ABB RAPID module: Module1_backup.mod

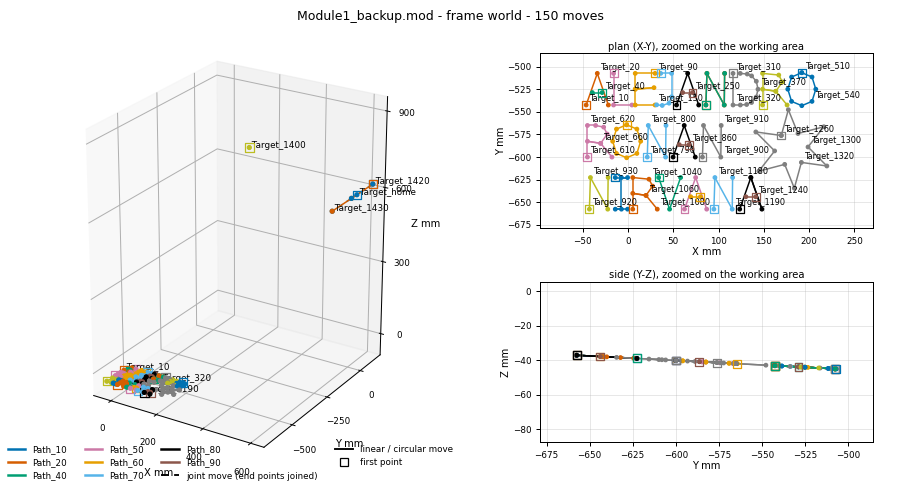
[picture p0: tool path of Module1_backup.mod in frame world, 150 of 178 moves have a stored position in this frame; points joined in program order, loops and branches not executed]
MODULE Module1
    PERS tooldata TOOLLAB1:=[TRUE,[[-6.48,-1.157,131.856],[0.965925826,0,0.258819045,0]],[1,[0,0,1],[1,0,0,0],0,0,0]];
    TASK PERS wobjdata Workobject_4:=[FALSE,TRUE,"",[[-82.07,-709.823595625,-134.482953476],[0.018509898,0.706864473,0.706864473,-0.018509898]],[[0,0,-100],[1,0,0,0]]];
    CONST robtarget Target_10:=[[162.356,35.679,0],[1,0,0,0],[-2,-1,0,1],[9E+09,9E+09,9E+09,9E+09,9E+09,9E+09]];
    CONST robtarget Target_20:=[[197.357,47.989,0],[1,0,0,0],[-2,-1,0,1],[9E+09,9E+09,9E+09,9E+09,9E+09,9E+09]];
    CONST robtarget Target_30:=[[162.356,60.2,0],[1,0,0,0],[-2,-1,0,1],[9E+09,9E+09,9E+09,9E+09,9E+09,9E+09]];
    CONST robtarget Target_40:=[[176.113,53.293,0],[1,0,0,0],[-2,-1,0,1],[9E+09,9E+09,9E+09,9E+09,9E+09,9E+09]];
    CONST robtarget Target_50:=[[176.113,42.487,0],[1,0,0,0],[-2,-1,0,1],[9E+09,9E+09,9E+09,9E+09,9E+09,9E+09]];
    VAR robtarget lift:=[[176.113,42.487,0],[0.707106781,0,0,-0.707106781],[-2,-1,0,1],[9E+09,9E+09,9E+09,9E+09,9E+09,9E+09]];
    CONST robtarget Target_60:=[[197.357,65.972,0],[1,0,0,0],[-2,-1,0,1],[9E+09,9E+09,9E+09,9E+09,9E+09,9E+09]];
    CONST robtarget Target_70:=[[162.356,65.972,0],[1,0,0,0],[-2,-1,0,1],[9E+09,9E+09,9E+09,9E+09,9E+09,9E+09]];
    CONST robtarget Target_80:=[[162.356,86.252,0],[1,0,0,0],[-2,-1,0,1],[9E+09,9E+09,9E+09,9E+09,9E+09,9E+09]];
    CONST robtarget Target_90:=[[197.357,111.808,0],[1,0,0,0],[-2,-1,0,1],[9E+09,9E+09,9E+09,9E+09,9E+09,9E+09]];
    CONST robtarget Target_100:=[[197.357,89.911,0],[1,0,0,0],[-2,-1,0,1],[9E+09,9E+09,9E+09,9E+09,9E+09,9E+09]];
    CONST robtarget Target_110:=[[179.857,89.911,0],[1,0,0,0],[-2,-1,0,1],[9E+09,9E+09,9E+09,9E+09,9E+09,9E+09]];
    CONST robtarget Target_120:=[[181.559,110.645,0],[1,0,0,0],[-2,-1,0,1],[9E+09,9E+09,9E+09,9E+09,9E+09,9E+09]];
    CONST robtarget Target_130:=[[179.857,89.911,0],[1,0,0,0],[-2,-1,0,1],[9E+09,9E+09,9E+09,9E+09,9E+09,9E+09]];
    CONST robtarget Target_140:=[[162.356,89.911,0],[1,0,0,0],[-2,-1,0,1],[9E+09,9E+09,9E+09,9E+09,9E+09,9E+09]];
    CONST robtarget Target_150:=[[162.356,111.808,0],[1,0,0,0],[-2,-1,0,1],[9E+09,9E+09,9E+09,9E+09,9E+09,9E+09]];
    CONST robtarget Target_160:=[[197.357,118.048,0],[1,0,0,0],[-2,-1,0,1],[9E+09,9E+09,9E+09,9E+09,9E+09,9E+09]];
    CONST robtarget Target_170:=[[197.357,130.103,0],[1,0,0,0],[-2,-1,0,1],[9E+09,9E+09,9E+09,9E+09,9E+09,9E+09]];
    CONST robtarget Target_180:=[[171.461,130.103,0],[1,0,0,0],[-2,-1,0,1],[9E+09,9E+09,9E+09,9E+09,9E+09,9E+09]];
    CONST robtarget Target_190:=[[164.37,127.295,0],[1,0,0,0],[-2,-1,0,1],[9E+09,9E+09,9E+09,9E+09,9E+09,9E+09]];
    CONST robtarget Target_200:=[[161.874,119.75,0],[1,0,0,0],[-2,-1,0,1],[9E+09,9E+09,9E+09,9E+09,9E+09,9E+09]];
    CONST robtarget Target_210:=[[162.555,113.567,0],[1,0,0,0],[-2,-1,0,1],[9E+09,9E+09,9E+09,9E+09,9E+09,9E+09]];
    CONST robtarget Target_220:=[[162.356,135.549,0],[1,0,0,0],[-2,-1,0,1],[9E+09,9E+09,9E+09,9E+09,9E+09,9E+09]];
    CONST robtarget Target_230:=[[197.357,147.859,0],[1,0,0,0],[-2,-1,0,1],[9E+09,9E+09,9E+09,9E+09,9E+09,9E+09]];
    CONST robtarget Target_240:=[[162.356,160.07,0],[1,0,0,0],[-2,-1,0,1],[9E+09,9E+09,9E+09,9E+09,9E+09,9E+09]];
    CONST robtarget Target_250:=[[176.113,153.163,0],[1,0,0,0],[-2,-1,0,1],[9E+09,9E+09,9E+09,9E+09,9E+09,9E+09]];
    CONST robtarget Target_260:=[[176.113,142.356,0],[1,0,0,0],[-2,-1,0,1],[9E+09,9E+09,9E+09,9E+09,9E+09,9E+09]];
    CONST robtarget Target_310:=[[197.357,197.978,0],[1,0,0,0],[-2,-1,0,1],[9E+09,9E+09,9E+09,9E+09,9E+09,9E+09]];
    CONST robtarget Target_320:=[[162.356,197.978,0],[1,0,0,0],[-2,-1,0,1],[9E+09,9E+09,9E+09,9E+09,9E+09,9E+09]];
    CONST robtarget Target_330:=[[162.356,206.033,0],[1,0,0,0],[-2,-1,0,1],[9E+09,9E+09,9E+09,9E+09,9E+09,9E+09]];
    CONST robtarget Target_340:=[[162.924,213.025,0],[1,0,0,0],[-2,-1,0,1],[9E+09,9E+09,9E+09,9E+09,9E+09,9E+09]];
    CONST robtarget Target_350:=[[165.164,218.429,0],[1,0,0,0],[-2,-1,0,1],[9E+09,9E+09,9E+09,9E+09,9E+09,9E+09]];
    CONST robtarget Target_360:=[[171.177,223.633,0],[1,0,0,0],[-2,-1,0,1],[9E+09,9E+09,9E+09,9E+09,9E+09,9E+09]];
    CONST robtarget Target_370:=[[179.829,225.576,0],[1,0,0,0],[-2,-1,0,1],[9E+09,9E+09,9E+09,9E+09,9E+09,9E+09]];
    CONST robtarget Target_380:=[[188.636,223.718,0],[1,0,0,0],[-2,-1,0,1],[9E+09,9E+09,9E+09,9E+09,9E+09,9E+09]];
    CONST robtarget Target_390:=[[194.578,218.485,0],[1,0,0,0],[-2,-1,0,1],[9E+09,9E+09,9E+09,9E+09,9E+09,9E+09]];
    CONST robtarget Target_400:=[[196.62,213.692,0],[1,0,0,0],[-2,-1,0,1],[9E+09,9E+09,9E+09,9E+09,9E+09,9E+09]];
    CONST robtarget Target_410:=[[197.357,205.948,0],[1,0,0,0],[-2,-1,0,1],[9E+09,9E+09,9E+09,9E+09,9E+09,9E+09]];
    CONST robtarget Target_420:=[[162.356,230.625,0],[1,0,0,0],[-2,-1,0,1],[9E+09,9E+09,9E+09,9E+09,9E+09,9E+09]];
    CONST robtarget Target_430:=[[197.357,230.625,0],[1,0,0,0],[-2,-1,0,1],[9E+09,9E+09,9E+09,9E+09,9E+09,9E+09]];
    CONST robtarget Target_450:=[[195.514,248.551,0],[1,0,0,0],[-2,-1,0,1],[9E+09,9E+09,9E+09,9E+09,9E+09,9E+09]];
    CONST robtarget Target_460:=[[187.856,252.522,0],[1,0,0,0],[-2,-1,0,1],[9E+09,9E+09,9E+09,9E+09,9E+09,9E+09]];
    CONST robtarget Target_470:=[[177.588,245.261,0],[1,0,0,0],[-2,-1,0,1],[9E+09,9E+09,9E+09,9E+09,9E+09,9E+09]];
    CONST robtarget Target_480:=[[179.857,230.625,0],[1,0,0,0],[-2,-1,0,1],[9E+09,9E+09,9E+09,9E+09,9E+09,9E+09]];
    CONST robtarget Target_490:=[[177.588,245.261,0],[1,0,0,0],[-2,-1,0,1],[9E+09,9E+09,9E+09,9E+09,9E+09,9E+09]];
    CONST robtarget Target_500:=[[162.356,257.713,0],[1,0,0,0],[-2,-1,0,1],[9E+09,9E+09,9E+09,9E+09,9E+09,9E+09]];
    CONST robtarget Target_510:=[[198.095,273.965,0],[1,0,0,0],[-2,-1,0,1],[9E+09,9E+09,9E+09,9E+09,9E+09,9E+09]];
    CONST robtarget Target_520:=[[193.358,285.254,0],[1,0,0,0],[-2,-1,0,1],[9E+09,9E+09,9E+09,9E+09,9E+09,9E+09]];
    CONST robtarget Target_530:=[[179.857,289.452,0],[1,0,0,0],[-2,-1,0,1],[9E+09,9E+09,9E+09,9E+09,9E+09,9E+09]];
    CONST robtarget Target_540:=[[166.384,285.254,0],[1,0,0,0],[-2,-1,0,1],[9E+09,9E+09,9E+09,9E+09,9E+09,9E+09]];
    CONST robtarget Target_550:=[[161.619,273.965,0],[1,0,0,0],[-2,-1,0,1],[9E+09,9E+09,9E+09,9E+09,9E+09,9E+09]];
    CONST robtarget Target_560:=[[166.384,262.676,0],[1,0,0,0],[-2,-1,0,1],[9E+09,9E+09,9E+09,9E+09,9E+09,9E+09]];
    CONST robtarget Target_570:=[[179.857,258.507,0],[1,0,0,0],[-2,-1,0,1],[9E+09,9E+09,9E+09,9E+09,9E+09,9E+09]];
    CONST robtarget Target_590:=[[193.358,262.705,0],[1,0,0,0],[-2,-1,0,1],[9E+09,9E+09,9E+09,9E+09,9E+09,9E+09]];
    CONST robtarget Target_600:=[[198.095,273.965,0],[1,0,0,0],[-2,-1,0,1],[9E+09,9E+09,9E+09,9E+09,9E+09,9E+09]];
    CONST robtarget Target_270:=[[162.356,168.011,0],[1,0,0,0],[-2,-1,0,1],[9E+09,9E+09,9E+09,9E+09,9E+09,9E+09]];
    CONST robtarget Target_280:=[[197.357,169.146,0],[1,0,0,0],[-2,-1,0,1],[9E+09,9E+09,9E+09,9E+09,9E+09,9E+09]];
    CONST robtarget Target_290:=[[162.356,188.278,0],[1,0,0,0],[-2,-1,0,1],[9E+09,9E+09,9E+09,9E+09,9E+09,9E+09]];
    CONST robtarget Target_300:=[[197.357,188.717,0],[1,0,0,0],[-2,-1,0,1],[9E+09,9E+09,9E+09,9E+09,9E+09,9E+09]];
    CONST robtarget Target_610:=[[104.728,37.097,0],[1,0,0,0],[-2,-1,0,1],[9E+09,9E+09,9E+09,9E+09,9E+09,9E+09]];
    CONST robtarget Target_620:=[[139.729,37.097,0],[1,0,0,0],[-2,-1,0,1],[9E+09,9E+09,9E+09,9E+09,9E+09,9E+09]];
    CONST robtarget Target_630:=[[139.729,46.117,0],[1,0,0,0],[-2,-1,0,1],[9E+09,9E+09,9E+09,9E+09,9E+09,9E+09]];
    CONST robtarget Target_640:=[[137.885,55.023,0],[1,0,0,0],[-2,-1,0,1],[9E+09,9E+09,9E+09,9E+09,9E+09,9E+09]];
    CONST robtarget Target_650:=[[130.227,58.994,0],[1,0,0,0],[-2,-1,0,1],[9E+09,9E+09,9E+09,9E+09,9E+09,9E+09]];
    CONST robtarget Target_660:=[[119.959,51.733,0],[1,0,0,0],[-2,-1,0,1],[9E+09,9E+09,9E+09,9E+09,9E+09,9E+09]];
    CONST robtarget Target_670:=[[122.228,37.097,0],[1,0,0,0],[-2,-1,0,1],[9E+09,9E+09,9E+09,9E+09,9E+09,9E+09]];
    CONST robtarget Target_680:=[[119.959,51.733,0],[1,0,0,0],[-2,-1,0,1],[9E+09,9E+09,9E+09,9E+09,9E+09,9E+09]];
    CONST robtarget Target_690:=[[104.728,64.185,0],[1,0,0,0],[-2,-1,0,1],[9E+09,9E+09,9E+09,9E+09,9E+09,9E+09]];
    CONST robtarget Target_700:=[[140.466,80.438,0],[1,0,0,0],[-2,-1,0,1],[9E+09,9E+09,9E+09,9E+09,9E+09,9E+09]];
    CONST robtarget Target_710:=[[135.73,91.726,0],[1,0,0,0],[-2,-1,0,1],[9E+09,9E+09,9E+09,9E+09,9E+09,9E+09]];
    CONST robtarget Target_720:=[[122.228,95.924,0],[1,0,0,0],[-2,-1,0,1],[9E+09,9E+09,9E+09,9E+09,9E+09,9E+09]];
    CONST robtarget Target_730:=[[108.755,91.726,0],[1,0,0,0],[-2,-1,0,1],[9E+09,9E+09,9E+09,9E+09,9E+09,9E+09]];
    CONST robtarget Target_740:=[[103.99,80.438,0],[1,0,0,0],[-2,-1,0,1],[9E+09,9E+09,9E+09,9E+09,9E+09,9E+09]];
    CONST robtarget Target_750:=[[108.755,69.149,0],[1,0,0,0],[-2,-1,0,1],[9E+09,9E+09,9E+09,9E+09,9E+09,9E+09]];
    CONST robtarget Target_760:=[[122.228,64.979,0],[1,0,0,0],[-2,-1,0,1],[9E+09,9E+09,9E+09,9E+09,9E+09,9E+09]];
    CONST robtarget Target_770:=[[135.73,69.177,0],[1,0,0,0],[-2,-1,0,1],[9E+09,9E+09,9E+09,9E+09,9E+09,9E+09]];
    CONST robtarget Target_780:=[[140.466,80.438,0],[1,0,0,0],[-2,-1,0,1],[9E+09,9E+09,9E+09,9E+09,9E+09,9E+09]];
    CONST robtarget Target_790:=[[104.728,103.2,0],[1,0,0,0],[-2,-1,0,1],[9E+09,9E+09,9E+09,9E+09,9E+09,9E+09]];
    CONST robtarget Target_800:=[[139.729,104.334,0],[1,0,0,0],[-2,-1,0,1],[9E+09,9E+09,9E+09,9E+09,9E+09,9E+09]];
    CONST robtarget Target_810:=[[104.728,123.466,0],[1,0,0,0],[-2,-1,0,1],[9E+09,9E+09,9E+09,9E+09,9E+09,9E+09]];
    CONST robtarget Target_820:=[[139.729,123.905,0],[1,0,0,0],[-2,-1,0,1],[9E+09,9E+09,9E+09,9E+09,9E+09,9E+09]];
    CONST robtarget Target_830:=[[104.728,131.748,0],[1,0,0,0],[-2,-1,0,1],[9E+09,9E+09,9E+09,9E+09,9E+09,9E+09]];
    CONST robtarget Target_840:=[[139.729,144.058,0],[1,0,0,0],[-2,-1,0,1],[9E+09,9E+09,9E+09,9E+09,9E+09,9E+09]];
    CONST robtarget Target_850:=[[104.728,156.269,0],[1,0,0,0],[-2,-1,0,1],[9E+09,9E+09,9E+09,9E+09,9E+09,9E+09]];
    CONST robtarget Target_860:=[[118.484,149.362,0],[1,0,0,0],[-2,-1,0,1],[9E+09,9E+09,9E+09,9E+09,9E+09,9E+09]];
    CONST robtarget Target_870:=[[118.484,138.555,0],[1,0,0,0],[-2,-1,0,1],[9E+09,9E+09,9E+09,9E+09,9E+09,9E+09]];
    CONST robtarget Target_880:=[[104.728,164.211,0],[1,0,0,0],[-2,-1,0,1],[9E+09,9E+09,9E+09,9E+09,9E+09,9E+09]];
    CONST robtarget Target_890:=[[139.729,165.345,0],[1,0,0,0],[-2,-1,0,1],[9E+09,9E+09,9E+09,9E+09,9E+09,9E+09]];
    CONST robtarget Target_900:=[[104.728,184.477,0],[1,0,0,0],[-2,-1,0,1],[9E+09,9E+09,9E+09,9E+09,9E+09,9E+09]];
    CONST robtarget Target_910:=[[139.729,184.916,0],[1,0,0,0],[-2,-1,0,1],[9E+09,9E+09,9E+09,9E+09,9E+09,9E+09]];
    CONST robtarget Target_920:=[[47.099,39.267,0],[1,0,0,0],[-2,-1,0,1],[9E+09,9E+09,9E+09,9E+09,9E+09,9E+09]];
    CONST robtarget Target_930:=[[82.1,40.402,0],[1,0,0,0],[-2,-1,0,1],[9E+09,9E+09,9E+09,9E+09,9E+09,9E+09]];
    CONST robtarget Target_940:=[[47.099,59.533,0],[1,0,0,0],[-2,-1,0,1],[9E+09,9E+09,9E+09,9E+09,9E+09,9E+09]];
    CONST robtarget Target_950:=[[82.1,59.973,0],[1,0,0,0],[-2,-1,0,1],[9E+09,9E+09,9E+09,9E+09,9E+09,9E+09]];
    CONST robtarget Target_960:=[[82.1,67.872,0],[1,0,0,0],[-2,-1,0,1],[9E+09,9E+09,9E+09,9E+09,9E+09,9E+09]];
    CONST robtarget Target_970:=[[82.1,81.43,0],[1,0,0,0],[-2,-1,0,1],[9E+09,9E+09,9E+09,9E+09,9E+09,9E+09]];
    CONST robtarget Target_980:=[[82.1,74.651,0],[1,0,0,0],[-2,-1,0,1],[9E+09,9E+09,9E+09,9E+09,9E+09,9E+09]];
    CONST robtarget Target_990:=[[47.099,74.651,0],[1,0,0,0],[-2,-1,0,1],[9E+09,9E+09,9E+09,9E+09,9E+09,9E+09]];
    CONST robtarget Target_1000:=[[47.099,67.872,0],[1,0,0,0],[-2,-1,0,1],[9E+09,9E+09,9E+09,9E+09,9E+09,9E+09]];
    CONST robtarget Target_1010:=[[47.099,81.43,0],[1,0,0,0],[-2,-1,0,1],[9E+09,9E+09,9E+09,9E+09,9E+09,9E+09]];
    CONST robtarget Target_1020:=[[47.099,87.188,0],[1,0,0,0],[-2,-1,0,1],[9E+09,9E+09,9E+09,9E+09,9E+09,9E+09]];
    CONST robtarget Target_1030:=[[82.1,87.188,0],[1,0,0,0],[-2,-1,0,1],[9E+09,9E+09,9E+09,9E+09,9E+09,9E+09]];
    CONST robtarget Target_1040:=[[80.257,105.114,0],[1,0,0,0],[-2,-1,0,1],[9E+09,9E+09,9E+09,9E+09,9E+09,9E+09]];
    CONST robtarget Target_1050:=[[72.598,109.085,0],[1,0,0,0],[-2,-1,0,1],[9E+09,9E+09,9E+09,9E+09,9E+09,9E+09]];
    CONST robtarget Target_1060:=[[62.331,101.824,0],[1,0,0,0],[-2,-1,0,1],[9E+09,9E+09,9E+09,9E+09,9E+09,9E+09]];
    CONST robtarget Target_1070:=[[64.6,87.188,0],[1,0,0,0],[-2,-1,0,1],[9E+09,9E+09,9E+09,9E+09,9E+09,9E+09]];
    CONST robtarget Target_1075:=[[62.331,101.824,0],[1,0,0,0],[-2,-1,0,1],[9E+09,9E+09,9E+09,9E+09,9E+09,9E+09]];
    CONST robtarget Target_1080:=[[47.099,114.276,0],[1,0,0,0],[-2,-1,0,1],[9E+09,9E+09,9E+09,9E+09,9E+09,9E+09]];
    CONST robtarget Target_1090:=[[82.1,115.808,0],[1,0,0,0],[-2,-1,0,1],[9E+09,9E+09,9E+09,9E+09,9E+09,9E+09]];
    CONST robtarget Target_1100:=[[47.099,127.876,0],[1,0,0,0],[-2,-1,0,1],[9E+09,9E+09,9E+09,9E+09,9E+09,9E+09]];
    CONST robtarget Target_1110:=[[82.1,140.073,0],[1,0,0,0],[-2,-1,0,1],[9E+09,9E+09,9E+09,9E+09,9E+09,9E+09]];
    CONST robtarget Target_1120:=[[47.099,144.37,0],[1,0,0,0],[-2,-1,0,1],[9E+09,9E+09,9E+09,9E+09,9E+09,9E+09]];
    CONST robtarget Target_1130:=[[82.1,156.68,0],[1,0,0,0],[-2,-1,0,1],[9E+09,9E+09,9E+09,9E+09,9E+09,9E+09]];
    CONST robtarget Target_1140:=[[47.099,168.891,0],[1,0,0,0],[-2,-1,0,1],[9E+09,9E+09,9E+09,9E+09,9E+09,9E+09]];
    CONST robtarget Target_1150:=[[60.856,161.984,0],[1,0,0,0],[-2,-1,0,1],[9E+09,9E+09,9E+09,9E+09,9E+09,9E+09]];
    CONST robtarget Target_1160:=[[60.856,151.177,0],[1,0,0,0],[-2,-1,0,1],[9E+09,9E+09,9E+09,9E+09,9E+09,9E+09]];
    CONST robtarget Target_1170:=[[47.099,176.833,0],[1,0,0,0],[-2,-1,0,1],[9E+09,9E+09,9E+09,9E+09,9E+09,9E+09]];
    CONST robtarget Target_1180:=[[82.1,177.967,0],[1,0,0,0],[-2,-1,0,1],[9E+09,9E+09,9E+09,9E+09,9E+09,9E+09]];
    CONST robtarget Target_1190:=[[47.099,197.099,0],[1,0,0,0],[-2,-1,0,1],[9E+09,9E+09,9E+09,9E+09,9E+09,9E+09]];
    CONST robtarget Target_1200:=[[82.1,197.538,0],[1,0,0,0],[-2,-1,0,1],[9E+09,9E+09,9E+09,9E+09,9E+09,9E+09]];
    CONST robtarget Target_1210:=[[47.099,205.381,0],[1,0,0,0],[-2,-1,0,1],[9E+09,9E+09,9E+09,9E+09,9E+09,9E+09]];
    CONST robtarget Target_1220:=[[82.1,217.691,0],[1,0,0,0],[-2,-1,0,1],[9E+09,9E+09,9E+09,9E+09,9E+09,9E+09]];
    CONST robtarget Target_1230:=[[47.099,229.902,0],[1,0,0,0],[-2,-1,0,1],[9E+09,9E+09,9E+09,9E+09,9E+09,9E+09]];
    CONST robtarget Target_1240:=[[60.856,222.995,0],[1,0,0,0],[-2,-1,0,1],[9E+09,9E+09,9E+09,9E+09,9E+09,9E+09]];
    CONST robtarget Target_1250:=[[60.856,212.188,0],[1,0,0,0],[-2,-1,0,1],[9E+09,9E+09,9E+09,9E+09,9E+09,9E+09]];
    CONST robtarget Target_1260:=[[128.621,251.308,0],[1,0,0,0],[-2,-1,0,1],[9E+09,9E+09,9E+09,9E+09,9E+09,9E+09]];
    CONST robtarget Target_1270:=[[157.133,259.115,0],[1,0,0,0],[-2,-1,0,1],[9E+09,9E+09,9E+09,9E+09,9E+09,9E+09]];
    CONST robtarget Target_1280:=[[130.799,269.761,0],[1,0,0,0],[-2,-1,0,1],[9E+09,9E+09,9E+09,9E+09,9E+09,9E+09]];
    CONST robtarget Target_1290:=[[138.293,298.357,0],[1,0,0,0],[-2,-1,0,1],[9E+09,9E+09,9E+09,9E+09,9E+09,9E+09]];
    CONST robtarget Target_1300:=[[115.907,280.874,0],[1,0,0,0],[-2,-1,0,1],[9E+09,9E+09,9E+09,9E+09,9E+09,9E+09]];
    CONST robtarget Target_1310:=[[94.89,301.662,0],[1,0,0,0],[-2,-1,0,1],[9E+09,9E+09,9E+09,9E+09,9E+09,9E+09]];
    CONST robtarget Target_1320:=[[98.837,273.533,0],[1,0,0,0],[-2,-1,0,1],[9E+09,9E+09,9E+09,9E+09,9E+09,9E+09]];
    CONST robtarget Target_1330:=[[70.325,265.726,0],[1,0,0,0],[-2,-1,0,1],[9E+09,9E+09,9E+09,9E+09,9E+09,9E+09]];
    CONST robtarget Target_1340:=[[96.659,255.08,0],[1,0,0,0],[-2,-1,0,1],[9E+09,9E+09,9E+09,9E+09,9E+09,9E+09]];
    CONST robtarget Target_1350:=[[89.164,226.485,0],[1,0,0,0],[-2,-1,0,1],[9E+09,9E+09,9E+09,9E+09,9E+09,9E+09]];
    CONST robtarget Target_1360:=[[111.551,243.968,0],[1,0,0,0],[-2,-1,0,1],[9E+09,9E+09,9E+09,9E+09,9E+09,9E+09]];
    CONST robtarget Target_1370:=[[132.568,223.179,0],[1,0,0,0],[-2,-1,0,1],[9E+09,9E+09,9E+09,9E+09,9E+09,9E+09]];
    CONST robtarget Target_1380:=[[128.621,251.308,0],[1,0,0,0],[-2,-1,0,1],[9E+09,9E+09,9E+09,9E+09,9E+09,9E+09]];
    CONST robtarget Target_1400:=[[436.026984813,-441.348230806,910.76900576],[0.642444421,0.276181237,0.662820128,-0.267691179],[-1,0,-1,1],[9E+09,9E+09,9E+09,9E+09,9E+09,9E+09]];
    CONST robtarget Target_1420:=[[623.722328095,118.842990746,619.183756173],[0.258818958,-0.000000006,0.96592585,-0.000000022],[0,-1,0,0],[9E+09,9E+09,9E+09,9E+09,9E+09,9E+09]];
    CONST robtarget Target_1440:=[[623.72233089,-41.157009755,619.183762427],[0.258818973,0.000000002,0.965925846,-0.000000006],[-1,0,-1,0],[9E+09,9E+09,9E+09,9E+09,9E+09,9E+09]];
    CONST robtarget Target_1430:=[[623.722326179,-181.156992829,619.183758277],[0.258818962,-0.000000009,0.965925849,0.000000006],[-1,0,-1,0],[9E+09,9E+09,9E+09,9E+09,9E+09,9E+09]];
    CONST robtarget Target_home:=[[623.722296887,-1.157,619.183844617],[0.258819045,0,0.965925826,0],[-1,0,-1,0],[9E+09,9E+09,9E+09,9E+09,9E+09,9E+09]];




    PROC main()
        WHILE TRUE DO
            Reset DO_01;
            Reset DO_02;
            Reset DO_03;
            Reset FWD_Conveyor;
            Reset BWD_Conveyor;
            IF DI_01=1 THEN
                Move_banda_fwd;
                Path_10;
                Rutina_dibujo;
                Path_10;
                Move_banda_fwd;
            ENDIF
            IF DI_02=1 THEN
                SET DO_02;
                Path_Man;
                RESET DO_02;
            ENDIF
            IF DI_03=1 THEN
                SET DO_03;
                Path_10;
                Path_Aura;
                Path_Aura;
                Path_Aura;
                Path_10;
                RESET DO_03;
            ENDIF
        ENDWHILE
!        Path_10;
!        Rutina_dibujo;
!        Path_10;
    ENDPROC

    PROC Move_banda_fwd()
        Set FWD_conveyor;
        SET BWD_Conveyor;
        WaitTime 2.5 ;
        Reset BWD_conveyor;
        WaitTime 1 ;
    ENDPROC
    PROC Move_banda_bwd()
        RESET FWD_Conveyor;
        Set BWD_conveyor;
        WaitTime 2.5 ;
        RESET BWD_conveyor;
        WaitTime 1 ;
    ENDPROC

    PROC Rutina_dibujo()
        Path_20;
        Path_40;
        Path_50;
        Path_60;
        Path_70;
        Path_80;
        Path_90;
        Path_95;
        Path_100;
        Path_110;
        Path_120;
        Path_130;
        Path_140;
        Path_150;
        Path_160;
        Path_170;
        Path_180;
        Path_190;
        Path_200;
        Path_210;
        Path_220;
        Path_230;
        Path_240;
        Path_250;
        Path_260;
        Path_270;
        Path_280;
        Path_290;
    ENDPROC

    PROC Path_10()
        MoveJ Target_home,v150,z1,TOOLLAB1\WObj:=wobj0;
    ENDPROC
    PROC Path_20()
        MoveJ Target_10,v300,z1,TOOLLAB1\WObj:=Workobject_4;
        MoveL Target_20,v300,z1,TOOLLAB1\WObj:=Workobject_4;
        MoveL Target_30,v300,z1,TOOLLAB1\WObj:=Workobject_4;
        lift := Offs(Target_30, 0, 0, -50);
        MoveJ lift,v300,z1,TOOLLAB1\WObj:=Workobject_4;
    ENDPROC



    PROC Path_40()
        MoveJ Target_40,v300,z1,TOOLLAB1\WObj:=Workobject_4;
        MoveL Target_50,v300,z1,TOOLLAB1\WObj:=Workobject_4;
        lift := Offs(Target_50, 0, 0, -50);
        MoveJ lift,v300,z1,TOOLLAB1\WObj:=Workobject_4;
    ENDPROC

    PROC Path_50()
        MoveJ Target_60,v300,z1,TOOLLAB1\WObj:=Workobject_4;
        MoveL Target_70,v300,z1,TOOLLAB1\WObj:=Workobject_4;
        MoveL Target_80,v300,z1,TOOLLAB1\WObj:=Workobject_4;
        lift := Offs(Target_80, 0, 0, -50);
        MoveJ lift,v300,z1,TOOLLAB1\WObj:=Workobject_4;
    ENDPROC
    PROC Path_60()
        MoveJ Target_90,v300,z1,TOOLLAB1\WObj:=Workobject_4;
        MoveL Target_100,v300,z1,TOOLLAB1\WObj:=Workobject_4;
        MoveL Target_110,v300,z1,TOOLLAB1\WObj:=Workobject_4;
        MoveL Target_120,v300,z1,TOOLLAB1\WObj:=Workobject_4;
        MoveL Target_130,v300,z1,TOOLLAB1\WObj:=Workobject_4;
        MoveL Target_140,v300,z1,TOOLLAB1\WObj:=Workobject_4;
        MoveL Target_150,v300,z1,TOOLLAB1\WObj:=Workobject_4;
        lift := Offs(Target_150, 0, 0, -50);
        MoveJ lift,v300,z1,TOOLLAB1\WObj:=Workobject_4;
    ENDPROC
    PROC Path_70()
        MoveJ Target_160,v300,z1,TOOLLAB1\WObj:=Workobject_4;
        MoveL Target_170,v300,z1,TOOLLAB1\WObj:=Workobject_4;
        MoveL Target_180,v300,z1,TOOLLAB1\WObj:=Workobject_4;
        MoveL Target_190,v300,z1,TOOLLAB1\WObj:=Workobject_4;
        MoveL Target_200,v300,z1,TOOLLAB1\WObj:=Workobject_4;
        MoveL Target_210,v300,z1,TOOLLAB1\WObj:=Workobject_4;
        lift := Offs(Target_210, 0, 0, -50);
        MoveJ lift,v300,z1,TOOLLAB1\WObj:=Workobject_4;
    ENDPROC
    PROC Path_30()

    ENDPROC
    PROC Path_80()
        MoveJ Target_220,v300,z1,TOOLLAB1\WObj:=Workobject_4;
        MoveL Target_230,v300,z1,TOOLLAB1\WObj:=Workobject_4;
        MoveL Target_240,v300,z1,TOOLLAB1\WObj:=Workobject_4;
        lift := Offs(Target_240, 0, 0, -50);
        MoveJ lift,v300,z1,TOOLLAB1\WObj:=Workobject_4;
    ENDPROC
    PROC Path_90()
        MoveJ Target_250,v300,z1,TOOLLAB1\WObj:=Workobject_4;
        MoveL Target_260,v300,z1,TOOLLAB1\WObj:=Workobject_4;
        lift := Offs(Target_260, 0, 0, -50);
        MoveJ lift,v300,z1,TOOLLAB1\WObj:=Workobject_4;
    ENDPROC
    PROC Path_100()
        MoveJ Target_310,v300,z1,TOOLLAB1\WObj:=Workobject_4;
        MoveL Target_320,v300,z1,TOOLLAB1\WObj:=Workobject_4;
        MoveL Target_330,v300,z1,TOOLLAB1\WObj:=Workobject_4;
        MoveL Target_340,v300,z1,TOOLLAB1\WObj:=Workobject_4;
        MoveL Target_350,v300,z1,TOOLLAB1\WObj:=Workobject_4;
        MoveL Target_360,v300,z1,TOOLLAB1\WObj:=Workobject_4;
        MoveL Target_370,v300,z1,TOOLLAB1\WObj:=Workobject_4;
        MoveL Target_380,v300,z1,TOOLLAB1\WObj:=Workobject_4;
        MoveL Target_390,v300,z1,TOOLLAB1\WObj:=Workobject_4;
        MoveL Target_400,v300,z1,TOOLLAB1\WObj:=Workobject_4;
        MoveL Target_410,v300,z1,TOOLLAB1\WObj:=Workobject_4;
        lift := Offs(Target_410, 0, 0, -50);
        MoveJ lift,v300,z1,TOOLLAB1\WObj:=Workobject_4;
    ENDPROC
    PROC Path_110()
        MoveJ Target_420,v300,z1,TOOLLAB1\WObj:=Workobject_4;
        MoveL Target_430,v300,z1,TOOLLAB1\WObj:=Workobject_4;
        MoveL Target_450,v300,z1,TOOLLAB1\WObj:=Workobject_4;
        MoveL Target_460,v300,z1,TOOLLAB1\WObj:=Workobject_4;
        MoveL Target_470,v300,z1,TOOLLAB1\WObj:=Workobject_4;
        MoveL Target_480,v300,z1,TOOLLAB1\WObj:=Workobject_4;
        MoveL Target_490,v300,z1,TOOLLAB1\WObj:=Workobject_4;
        MoveL Target_500,v300,z1,TOOLLAB1\WObj:=Workobject_4;
        lift := Offs(Target_500, 0, 0, -50);
        MoveJ lift,v300,z1,TOOLLAB1\WObj:=Workobject_4;
    ENDPROC
    PROC Path_120()
        MoveJ Target_510,v300,z1,TOOLLAB1\WObj:=Workobject_4;
        MoveL Target_520,v300,z1,TOOLLAB1\WObj:=Workobject_4;
        MoveL Target_530,v300,z1,TOOLLAB1\WObj:=Workobject_4;
        MoveL Target_540,v300,z1,TOOLLAB1\WObj:=Workobject_4;
        MoveL Target_550,v300,z1,TOOLLAB1\WObj:=Workobject_4;
        MoveL Target_560,v300,z1,TOOLLAB1\WObj:=Workobject_4;
        MoveL Target_570,v300,z1,TOOLLAB1\WObj:=Workobject_4;
        MoveL Target_590,v300,z1,TOOLLAB1\WObj:=Workobject_4;
        MoveL Target_600,v300,z1,TOOLLAB1\WObj:=Workobject_4;
        lift := Offs(Target_210, 0, 0, -50);
        MoveJ lift,v300,z1,TOOLLAB1\WObj:=Workobject_4;
    ENDPROC
    PROC Path_95()
        MoveJ Target_270,v300,z1,TOOLLAB1\WObj:=Workobject_4;
        MoveL Target_280,v300,z1,TOOLLAB1\WObj:=Workobject_4;
        MoveL Target_290,v300,z1,TOOLLAB1\WObj:=Workobject_4;
        MoveL Target_300,v300,z1,TOOLLAB1\WObj:=Workobject_4;
        lift := Offs(Target_300, 0, 0, -50);
        MoveJ lift,v300,z1,TOOLLAB1\WObj:=Workobject_4;
    ENDPROC
    PROC Path_85()
        MoveJ Target_270,v300,z1,TOOLLAB1\WObj:=Workobject_4;
        MoveL Target_280,v300,z1,TOOLLAB1\WObj:=Workobject_4;
        MoveL Target_290,v300,z1,TOOLLAB1\WObj:=Workobject_4;
        MoveL Target_300,v300,z1,TOOLLAB1\WObj:=Workobject_4;
        lift := Offs(Target_300, 0, 0, -50);
        MoveJ lift,v300,z1,TOOLLAB1\WObj:=Workobject_4;
    ENDPROC
    PROC Path_130()
        MoveJ Target_610,v300,z1,TOOLLAB1\WObj:=Workobject_4;
        MoveL Target_620,v300,z1,TOOLLAB1\WObj:=Workobject_4;
        MoveL Target_630,v300,z1,TOOLLAB1\WObj:=Workobject_4;
        MoveL Target_640,v300,z1,TOOLLAB1\WObj:=Workobject_4;
        MoveL Target_650,v300,z1,TOOLLAB1\WObj:=Workobject_4;
        MoveL Target_660,v300,z1,TOOLLAB1\WObj:=Workobject_4;
        MoveL Target_670,v300,z1,TOOLLAB1\WObj:=Workobject_4;
        MoveL Target_680,v300,z1,TOOLLAB1\WObj:=Workobject_4;
        MoveL Target_690,v300,z1,TOOLLAB1\WObj:=Workobject_4;
        lift := Offs(Target_690, 0, 0, -50);
        MoveJ lift,v300,z1,TOOLLAB1\WObj:=Workobject_4;
    ENDPROC
    PROC Path_140()
        MoveJ Target_700,v300,z1,TOOLLAB1\WObj:=Workobject_4;
        MoveL Target_710,v300,z1,TOOLLAB1\WObj:=Workobject_4;
        MoveL Target_720,v300,z1,TOOLLAB1\WObj:=Workobject_4;
        MoveL Target_730,v300,z1,TOOLLAB1\WObj:=Workobject_4;
        MoveL Target_740,v300,z1,TOOLLAB1\WObj:=Workobject_4;
        MoveL Target_750,v300,z1,TOOLLAB1\WObj:=Workobject_4;
        MoveL Target_760,v300,z1,TOOLLAB1\WObj:=Workobject_4;
        MoveL Target_770,v300,z1,TOOLLAB1\WObj:=Workobject_4;
        MoveL Target_780,v300,z1,TOOLLAB1\WObj:=Workobject_4;
        lift := Offs(Target_780, 0, 0, -50);
        MoveJ lift,v300,z1,TOOLLAB1\WObj:=Workobject_4;
    ENDPROC
    PROC Path_150()
        MoveJ Target_790,v300,z1,TOOLLAB1\WObj:=Workobject_4;
        MoveL Target_800,v300,z1,TOOLLAB1\WObj:=Workobject_4;
        MoveL Target_810,v300,z1,TOOLLAB1\WObj:=Workobject_4;
        MoveL Target_820,v300,z1,TOOLLAB1\WObj:=Workobject_4;
        lift := Offs(Target_820, 0, 0, -50);
        MoveJ lift,v300,z1,TOOLLAB1\WObj:=Workobject_4;
    ENDPROC
    PROC Path_160()
        MoveJ Target_830,v300,z1,TOOLLAB1\WObj:=Workobject_4;
        MoveL Target_840,v300,z1,TOOLLAB1\WObj:=Workobject_4;
        MoveL Target_850,v300,z1,TOOLLAB1\WObj:=Workobject_4;
        lift := Offs(Target_850, 0, 0, -50);
        MoveJ lift,v300,z1,TOOLLAB1\WObj:=Workobject_4;
    ENDPROC
    PROC Path_170()
        MoveJ Target_860,v300,z1,TOOLLAB1\WObj:=Workobject_4;
        MoveL Target_870,v300,z1,TOOLLAB1\WObj:=Workobject_4;
        lift := Offs(Target_870, 0, 0, -50);
        MoveJ lift,v300,z1,TOOLLAB1\WObj:=Workobject_4;
    ENDPROC
    PROC Path_180()
        MoveJ Target_880,v300,z1,TOOLLAB1\WObj:=Workobject_4;
        MoveL Target_890,v300,z1,TOOLLAB1\WObj:=Workobject_4;
        MoveL Target_900,v300,z1,TOOLLAB1\WObj:=Workobject_4;
        MoveL Target_910,v300,z1,TOOLLAB1\WObj:=Workobject_4;
        lift := Offs(Target_910, 0, 0, -50);
        MoveJ lift,v300,z1,TOOLLAB1\WObj:=Workobject_4;
    ENDPROC
    PROC Path_190()
        MoveJ Target_920,v300,z1,TOOLLAB1\WObj:=Workobject_4;
        MoveL Target_930,v300,z1,TOOLLAB1\WObj:=Workobject_4;
        MoveL Target_940,v300,z1,TOOLLAB1\WObj:=Workobject_4;
        MoveL Target_950,v300,z1,TOOLLAB1\WObj:=Workobject_4;
        lift := Offs(Target_950, 0, 0, -50);
        MoveJ lift,v300,z1,TOOLLAB1\WObj:=Workobject_4;
    ENDPROC
    PROC Path_200()
        MoveJ Target_960,v300,z1,TOOLLAB1\WObj:=Workobject_4;
        MoveL Target_970,v300,z1,TOOLLAB1\WObj:=Workobject_4;
        MoveL Target_980,v300,z1,TOOLLAB1\WObj:=Workobject_4;
        MoveL Target_990,v300,z1,TOOLLAB1\WObj:=Workobject_4;
        MoveL Target_1000,v300,z1,TOOLLAB1\WObj:=Workobject_4;
        MoveL Target_1010,v300,z1,TOOLLAB1\WObj:=Workobject_4;
        lift := Offs(Target_1010, 0, 0, -50);
        MoveJ lift,v300,z1,TOOLLAB1\WObj:=Workobject_4;
    ENDPROC
    PROC Path_210()
        MoveJ Target_1020,v300,z1,TOOLLAB1\WObj:=Workobject_4;
        MoveL Target_1030,v300,z1,TOOLLAB1\WObj:=Workobject_4;
        MoveL Target_1040,v300,z1,TOOLLAB1\WObj:=Workobject_4;
        MoveL Target_1050,v300,z1,TOOLLAB1\WObj:=Workobject_4;
        MoveL Target_1060,v300,z1,TOOLLAB1\WObj:=Workobject_4;
        MoveL Target_1070,v300,z1,TOOLLAB1\WObj:=Workobject_4;
        MoveL Target_1075,v300,z1,TOOLLAB1\WObj:=Workobject_4;
        MoveL Target_1080,v300,z1,TOOLLAB1\WObj:=Workobject_4;
        lift := Offs(Target_1080, 0, 0, -50);
        MoveJ lift,v300,z1,TOOLLAB1\WObj:=Workobject_4;
    ENDPROC
    PROC Path_220()
        MoveJ Target_1090,v300,z1,TOOLLAB1\WObj:=Workobject_4;
        MoveL Target_1100,v300,z1,TOOLLAB1\WObj:=Workobject_4;
        MoveL Target_1110,v300,z1,TOOLLAB1\WObj:=Workobject_4;
        lift := Offs(Target_1110, 0, 0, -50);
        MoveJ lift,v300,z1,TOOLLAB1\WObj:=Workobject_4;
    ENDPROC
    PROC Path_230()

    ENDPROC
    PROC Path_240()
        MoveJ Target_1120,v300,z1,TOOLLAB1\WObj:=Workobject_4;
        MoveL Target_1130,v300,z1,TOOLLAB1\WObj:=Workobject_4;
        MoveL Target_1140,v300,z1,TOOLLAB1\WObj:=Workobject_4;
        lift := Offs(Target_1140, 0, 0, -50);
        MoveJ lift,v300,z1,TOOLLAB1\WObj:=Workobject_4;
    ENDPROC
    PROC Path_250()
        MoveJ Target_1150,v300,z1,TOOLLAB1\WObj:=Workobject_4;
        MoveL Target_1160,v300,z1,TOOLLAB1\WObj:=Workobject_4;
        lift := Offs(Target_1160, 0, 0, -50);
        MoveJ lift,v300,z1,TOOLLAB1\WObj:=Workobject_4;
    ENDPROC
    PROC Path_260()
        MoveJ Target_1170,v300,z1,TOOLLAB1\WObj:=Workobject_4;
        MoveL Target_1180,v300,z1,TOOLLAB1\WObj:=Workobject_4;
        MoveL Target_1190,v300,z1,TOOLLAB1\WObj:=Workobject_4;
        MoveL Target_1200,v300,z1,TOOLLAB1\WObj:=Workobject_4;
        lift := Offs(Target_1200, 0, 0, -50);
        MoveJ lift,v300,z1,TOOLLAB1\WObj:=Workobject_4;
    ENDPROC
    PROC Path_270()
        MoveJ Target_1210,v300,z1,TOOLLAB1\WObj:=Workobject_4;
        MoveL Target_1220,v300,z1,TOOLLAB1\WObj:=Workobject_4;
        MoveL Target_1230,v300,z1,TOOLLAB1\WObj:=Workobject_4;
        MoveL Target_1220,v300,z1,TOOLLAB1\WObj:=Workobject_4;
        lift := Offs(Target_1220, 0, 0, -50);
        MoveJ lift,v300,z1,TOOLLAB1\WObj:=Workobject_4;
    ENDPROC
    PROC Path_280()
        MoveJ Target_1240,v300,z1,TOOLLAB1\WObj:=Workobject_4;
        MoveL Target_1250,v300,z1,TOOLLAB1\WObj:=Workobject_4;
        lift := Offs(Target_1250, 0, 0, -50);
        MoveJ lift,v300,z1,TOOLLAB1\WObj:=Workobject_4;
    ENDPROC
    PROC Path_290()
        MoveJ Target_1260,v300,z1,TOOLLAB1\WObj:=Workobject_4;
        MoveL Target_1270,v300,z1,TOOLLAB1\WObj:=Workobject_4;
        MoveL Target_1280,v300,z1,TOOLLAB1\WObj:=Workobject_4;
        MoveL Target_1290,v300,z1,TOOLLAB1\WObj:=Workobject_4;
        MoveL Target_1300,v300,z1,TOOLLAB1\WObj:=Workobject_4;
        MoveL Target_1310,v300,z1,TOOLLAB1\WObj:=Workobject_4;
        MoveL Target_1320,v300,z1,TOOLLAB1\WObj:=Workobject_4;
        MoveL Target_1330,v300,z1,TOOLLAB1\WObj:=Workobject_4;
        MoveL Target_1340,v300,z1,TOOLLAB1\WObj:=Workobject_4;
        MoveL Target_1350,v300,z1,TOOLLAB1\WObj:=Workobject_4;
        MoveL Target_1360,v300,z1,TOOLLAB1\WObj:=Workobject_4;
        MoveL Target_1370,v300,z1,TOOLLAB1\WObj:=Workobject_4;
        MoveL Target_1380,v300,z1,TOOLLAB1\WObj:=Workobject_4;
        lift := Offs(Target_1380, 0, 0, -50);
        MoveJ lift,v300,z1,TOOLLAB1\WObj:=Workobject_4;
    ENDPROC

    PROC Path_Man()
        MoveJ Target_1400,v100,z1,TOOLLAB1\WObj:=wobj0;
    ENDPROC


    PROC Path_Aura()
        MoveJ Target_1420,v300,z1,TOOLLAB1\WObj:=wobj0;
        MoveJ Target_1440,v300,z1,TOOLLAB1\WObj:=wobj0;
        MoveJ Target_1430,v300,z1,TOOLLAB1\WObj:=wobj0;
    ENDPROC
    PROC Path_320()
        MoveL Target_1420,v150,z1,TOOLLAB1\WObj:=wobj0;
        MoveL Target_1440,v150,z1,TOOLLAB1\WObj:=wobj0;
        MoveL Target_1430,v150,z1,TOOLLAB1\WObj:=wobj0;
    ENDPROC

ENDMODULE
